FUNCTION_BLOCK FB_PositionEncoder_1
(*
Position encoder resolution.

Constructor: 		Patryk Panylo
Company:		E. Riexinger GmbH
Date:			20.01.2014
Version:			1.00

Date:			Revision:		Who:				Comment
dd.mm.yyyy		x.xx			Initials			comment

*)
VAR_INPUT
	(* Enummerations *)
	
	(* Variables *)
	bEnable								:BOOL;							(* Enable FB *)

	dwEncCurrentValue					:DWORD;						(* Encoder current value [inc] *)

	stEncCfg								:ST_EncoderConfig;				(* Encoder configuration *)

	(* References *)

	(* Interfaces *)
	pAxis								:POINTER TO ST_AXIS_REF_V2;

	(* Instances *)
	fbActPosFilter							:FB_ValueFilter;					(* Actual position filter *)
END_VAR
VAR_OUTPUT
	(* Enummerations *)
	
	(* Variables *)

	(* References *)

	(* Interfaces *)

	(* Instances *)

END_VAR
VAR
	(* Enummerations *)

	(* Variables *)
	bFirstTime							:BOOL;							(* First cycle *)

	dwActPos							:DWORD;						(* Current position inc *)
	dwOldActPos							:DWORD;						(* Position old value *)
	dnPosDistance						:DINT;							(* Positon distance from encoder values *)
	dwPosOffset							:DWORD;						(* Positon offset from encoder values *)
	(* References *)
	lroffset:LREAL;
	(* Interfaces *)

	(* Instances *)
	fbVeloAccDecJerk					:FB_CalcVeloAccDecJerk;

END_VAR

IF NOT bEnable
THEN
	bFirstTime := FALSE;

	RETURN;
END_IF

IF NOT bFirstTime
THEN
	A_Init();

	bFirstTime := TRUE;
END_IF

A_GetPosition();
A_GetDynamics();

ACTION A_GetDynamics:

(* Current position value filtering *)
fbActPosFilter(
	bEnable := TRUE,
	lrInSignal := pAxis^.stPosition.lrActPos,
	lrDeltaMax := 0.001
);

(* Current dynamics *)
fbVeloAccDecJerk(
	bEnable := TRUE,
	bReset := FALSE,
	lrActPos := fbActPosFilter.lrOutSignal,
	lrSectorTime := pAxis^.stScaling.lrTaskCycle ,
	etDirection => pAxis^.stScaling.etDirection,
	lrCalcVelo => pAxis^.stDynamics.lrActVelo,
	bAccelerating => pAxis^.stAxisStates.bAccelerating,
	bDecelerating => pAxis^.stAxisStates.bDecelerating,
	lrCalcAcc => pAxis^.stDynamics.lrActAcc,
	lrCalcDec => pAxis^.stDynamics.lrActDec,
	lrCalcJerk => pAxis^.stDynamics.lrActJerk
);
END_ACTION

ACTION A_GetPosition:

dwActPos := dwEncCurrentValue;																			(* Current position inc *)

IF stEncCfg.etScalingMethod = ET_ScalingMethod_eSMRotary
THEN

	dnPosDistance := F_ModuloDistance(dwActPos, dwOldActPos, stEncCfg.dwModuloValue);						(* Position distance in inc *)

	dwActPos := dwActPos + DINT_TO_DWORD(dnPosDistance);												(* Current position in inc *)

	pAxis^.stPosition.dwActPos := dwActPos;																	(* Current position in inc *)

	pAxis^.stPosition.lrActPos := F_ConvertActPosResiduals(													(* Current position in technical units *)
		dwPos := dwActPos,
		pAxis := pAxis
	);

	pAxis^.stPosition.lrSetPos := F_ModR(pAxis^.stPosition.lrSetPos, stEncCfg.lrModuloFactor);						(* Current period positon in technical units *)

ELSIF stEncCfg.etScalingMethod = ET_ScalingMethod_eSMLinear
THEN

	(*IF stEncCfg.dwModuloValue > 0
	THEN

		dnPosDistance := DWORD_TO_DINT(dwActPos - dwOldActPos);											(* Position distance in inc *)

		IF dnPosDistance > (stEncCfg.dwModuloValue / 2)
		THEN
			dwPosOffset := dwPosOffset - stEncCfg.dwModuloValue;												(* Position offset in inc *)

		ELSIF dnPosDistance < -DWORD_TO_DINT(stEncCfg.dwModuloValue / 2)
		THEN
			dwPosOffset := dwPosOffset + stEncCfg.dwModuloValue;												(* Position offset in inc *)

		END_IF

		dwActPos := dwPosOffset + dwEncCurrentValue;														(* Current position in inc *)

	END_IF*)

	pAxis^.stPosition.dwActPos := dwActPos;																	(* Current position in inc *)

	pAxis^.stPosition.lrActPos := F_ConvertActPosResiduals(													(* Current position in technical units *)
								dwPos := dwActPos,
								pAxis := pAxis
							 );

END_IF

dwOldActPos := dwEncCurrentValue;

(*pAxis^.stPosition.lrActPos := pAxis^.stPosition.lrSetPos;*)														(* Current position in technical units *)
END_ACTION

ACTION A_Init:

dwOldActPos := dwEncCurrentValue;
END_ACTION

END_FUNCTION_BLOCK

(* stored: Version 1.1.0.1, ProductVersion 3.1.4024.15
   POU FB_PositionEncoder_1: Id {9256b2cd-7193-46f2-aee7-7123dd1f7b25}, SpecialFunc None
   Action A_GetDynamics: Id {51faffa5-eef8-44b3-ab43-cfa1c32f1924}
   Action A_GetPosition: Id {968c817d-2d29-4719-8ba4-3689a37963ee}
   Action A_Init: Id {6326c631-ddbe-44ad-b001-2d9646987617} *)
